(* Logix 5000 project; controller R400_500_XLS vendor 1 type 14 code 216 rev 31.11; software revision 31.01; part 10 of 32 *)
(* tags used below, declared in another part *)
   Alarm : SINT;   // Wait 3 seconds
   Cycles : UDT_CYCLE[11];
   DrnSmp : DINT;
   FC23_BaseConductivity : REAL;   // Base conductivity of the water prior to the injection
   Fill_Sump : DINT;
   M : DINT[5];   // Memory Bits
   MaxPressRecord : REAL;
   MinPressRecord : REAL;
   PureWaterTankFilling : BOOL;   // Start PWT filling
   Run : DINT;
   Service : DINT[2];   // Unused Service Mode Memory Bit
   Tmr : TIMER[107];
   WSH41_Hour : DINT;
   WSH41_Minute : DINT;
   WSH41_Second : DINT;
   abCycleDataToSCADA : BOOL[32];
   abInputToSCADA : BOOL[32];
   abOutputToSCADA : BOOL[32];
   aiCycleDataToSCADA : INT[16];
   AlarmTrigger : INT;   // Triggers the alarm screen if different of 0
   arAnalogInputToSCADA : REAL[8];
   arCycleDataToSCADA : REAL[8];
   bPureWaterFillingAuthorization : BOOL;   // Pure Water Filling Authorization Signal
   ChemCond : REAL;
   CR2Mode : SINT;   // 0= Cycle complete dry contact 1= External pure water valve
   CycleCounter : DINT;
   CyclePtr : DINT;   // Cycle Pointeur
   DryTemp : REAL;
   FinalRinseCond : REAL;
   I_Chm_1_Lvl_Sw : BOOL;   // Chemical Pump #1 level switch
   I_Chm_2_Lvl_Sw : BOOL;   // Chemical Pump #2 level switch
   I_Chm_3_Lvl_Sw : BOOL;   // Chemical Pump #3 level switch
   I_Chm_4_Lvl_Sw : BOOL;   // Chemical Pump #4 level switch
   I_Ld_Dr_Cls_Sw : BOOL;   // Load door close
   I_Ld_Dr_Obs_Sw : BOOL;   // Load door obstruction switch
   I_MCR : BOOL;   // MCR input
   I_Mtr_Ovrld : BOOL;   // Motor overload
   I_Pure_Water_Filling_Auth : BOOL;
   I_Pw_Tnk_Lvl_Sw : BOOL;   // Pure water tank level switch
   I_Pw_Tnk_Sft_Lvl_Sw : BOOL;   // Pure water tank safety level switch
   I_Shlf_Sw : BOOL;   // Shelf switch
   I_Smp_Lvl_Hgh : BOOL;   // Sump high level switch
   I_Smp_Lvl_Lw : BOOL;   // Sump low level switch
   I_Smp_Sft_Lvl_Sw : BOOL;   // Sump safety level switch
   I_Unld_Dr_Cls_Sw : BOOL;   // Unload door close
   I_Unld_Dr_Obs_Sw : BOOL;   // Unload door obstruction switch
   I_UnldDr_ClseSlnce_Bttn : BOOL;   // Door Close/ Silence button Unload Side
   I_UnldDr_Opn_Bttn : BOOL;   // Door Open button Unload side
   iAlarmToSCADA : INT;
   iSCADACycleCompleteTimeHr : INT;
   iSCADACycleCompleteTimeMin : INT;
   iSCADACycleCompleteTimeSec : INT;
   ONS_SCADA : INT;
   PmpPres : REAL;
   PureWaterTankFillingRequest : BOOL;
   PureWaterTankTemp : REAL;   // Pure water tank temperature
   Q_Adble_Alrm : BOOL;   // Audible Alarm and /Pilot Light: red connection
   Q_Chm_1 : BOOL;   // Chemical pump #1
   Q_Chm_2 : BOOL;   // Chemical pump #2
   Q_Chm_3 : BOOL;   // Chemical pump #3
   Q_Chm_4 : BOOL;   // Chemical pump #4
   Q_Cld_Wtr_Fll_Vlve : BOOL;   // Cold water sump fill valve
   Q_Cmmn_Alrm : BOOL;   // Dry contact For Alarm
   Q_Cndsr_Hflw_Vlve : BOOL;   // Condenser high flow cold water valve
   Q_Cndsr_Lflw_Vlve : BOOL;   // Condenser low flow cold water valve
   Q_Condensate_Return_Vlve : BOOL;   // Condensate Return CoolDown water valve
   Q_Cyc_Comp : BOOL;   // Dry Contact For Cycle Completed or Pure Water fill valve
   Q_Cyc_Run : BOOL;   // Pilot light: Green connection
   Q_Drn_Cldwn_Vlve : BOOL;   // Drain cool down water valve
   Q_Dry_Fan : BOOL;   // Vapor removal fan / Drying fan
   Q_Dry_Htr : BOOL;   // Drying heating elements
   Q_Dry_Iso_Vlve : BOOL;   // Drying Isolation Valve (Normally Closed Valve)
   Q_Ht_Rcvry_Tnk_Drn_Vlve : BOOL;   // Heat recovery tank drian valve
   Q_Ht_Wtr_Fll_Vlve : BOOL;   // Hot water sump fill valve
   Q_Int_Lght : BOOL;   // Interior Light
   Q_Ld_Dr_Clse_Vlv : BOOL;   // Load door close pilot valve
   Q_Ld_Dr_Opn_Vlv : BOOL;   // Load door open pilot valve
   Q_Pmp_Hgh_Spd : BOOL;   // Pump high speed
   Q_Pmp_Lw_Spd : BOOL;   // Pump low speed
   Q_Pure_Water_Filling_Request : BOOL;   // Pure Water Filling Request
   Q_Pw_Fll_Vlve : BOOL;   // Pure water sump/ Tank fill valve
   Q_Pw_Otlt_Vlve : BOOL;   // Pure water tank outlet valve
   Q_Pw_Tnk_Stm_Vlve : BOOL;   // PWT Steam Valve / Electric Heater
   Q_Smp_drn_Vlve : BOOL;   // Sump drain valve (Normally open valve)
   Q_Smp_Stm_Vlve : BOOL;   // Sump steam valve/ Electrical Heater
   Q_Trsfr_Vlve : BOOL;   // Transfer Valve (Normally Open Valve)
   Q_Unld_Dr_Clse_Vlve : BOOL;   // Unload door close pilot valve
   Q_Unld_Dr_Opn_Vlve : BOOL;   // Unload door open pilot valve
   rSCADACompensatedSetPoint : REAL;
   SumpTemp : REAL;   // Sump temperature in °C
   TreatmentPtr : DINT;
   udtPureWaterHandshakeFromSCADA : UDT_PORT_HANDSHAKE_FROM_SCADA;
   udtPureWaterHandshakeToSCADA : UDT_PORT_HANDSHAKE_TO_SCADA;
   Unit : Hrdwre;   // Unit Configuration
(* MainProgram, continued *)

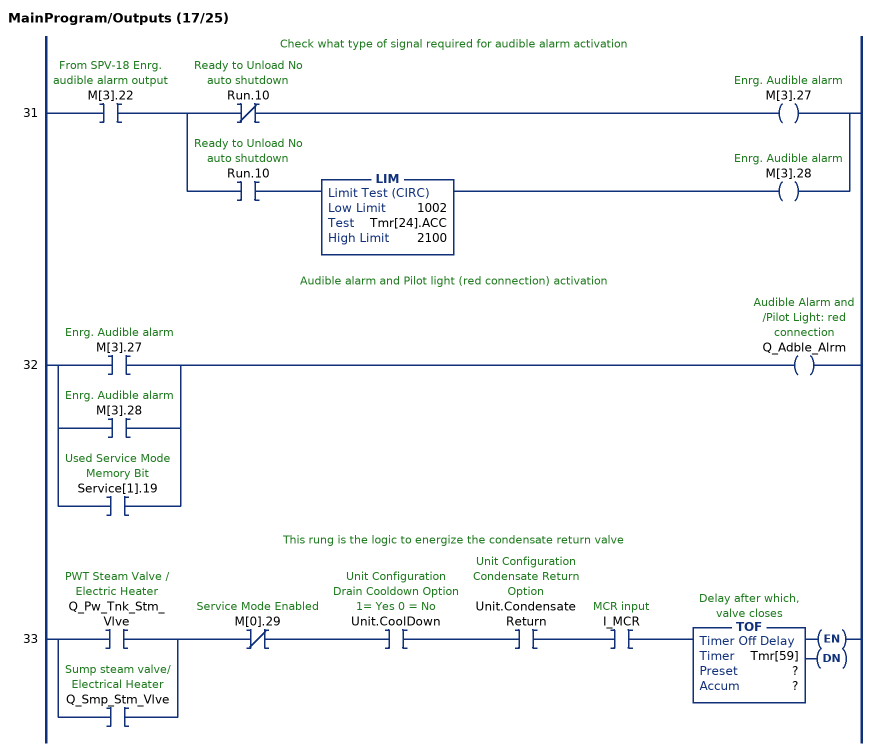
   [picture p153: MainProgram/Outputs rungs 31-33]
   // Check what type of signal required for audible alarm activation
   31: XIC(M[3].22)[XIO(Run.10) OTE(M[3].27) ,XIC(Run.10) LIM(1002,Tmr[24].ACC,2100) OTE(M[3].28) ];
   // Audible alarm and Pilot light (red connection) activation
   32: [XIC(M[3].27) ,XIC(M[3].28) ,XIC(Service[1].19) ]OTE(Q_Adble_Alrm);
   // This rung is the logic to energize the condensate return valve
   33: [XIC(Q_Pw_Tnk_Stm_Vlve) ,XIC(Q_Smp_Stm_Vlve) ]XIO(M[0].29)XIC(Unit.CoolDown)XIC(Unit.CondensateReturn)XIC(I_MCR)TOF(Tmr[59],?,?);
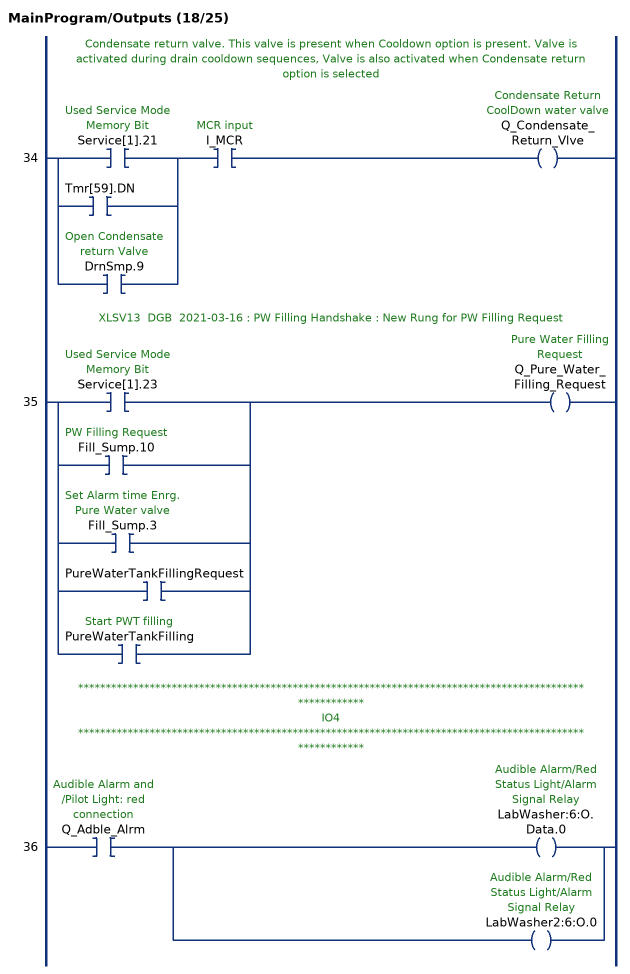
   // Condensate return valve. This valve is present when Cooldown option is present. Valve is activated during drain cooldown sequences, Valve is also activated when Condensate return option is selected
   34: [XIC(Service[1].21) ,XIC(Tmr[59].DN) ,XIC(DrnSmp.9) ]XIC(I_MCR)OTE(Q_Condensate_Return_Vlve);
   // XLSV13  DGB  2021-03-16 : PW Filling Handshake : New Rung for PW Filling Request
   35: [XIC(Service[1].23) ,XIC(Fill_Sump.10) ,XIC(Fill_Sump.3) ,XIC(PureWaterTankFillingRequest) ,XIC(PureWaterTankFilling) ]OTE(Q_Pure_Water_Filling_Request);
   // ********************************************************************************************************
   // IO4
   // ********************************************************************************************************
   36: XIC(Q_Adble_Alrm)[OTE(LabWasher:6:O.Data.0) ,OTE(LabWasher2:6:O.0) ];
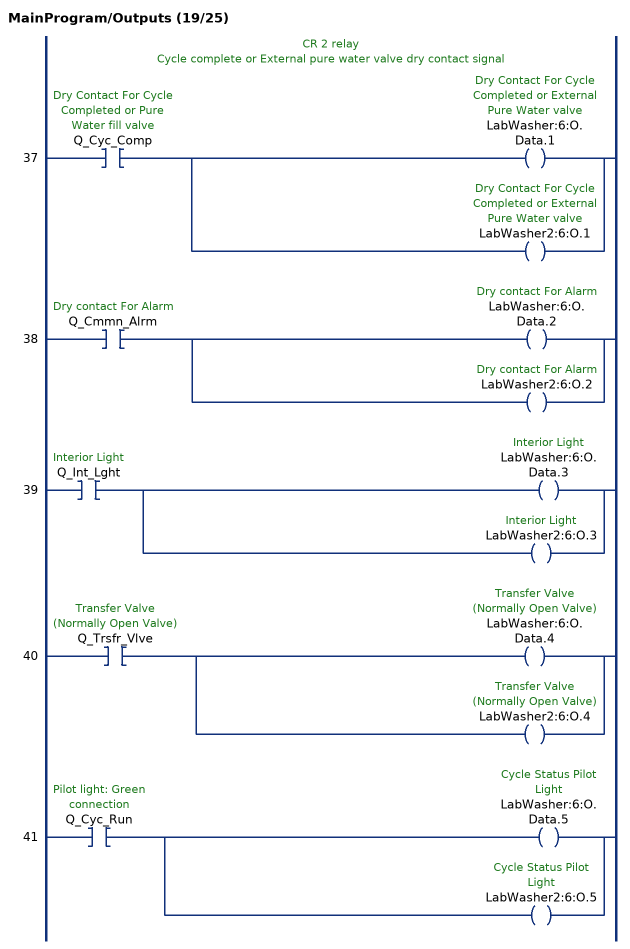
   // CR 2 relay
   // Cycle complete or External pure water valve dry contact signal
   37: XIC(Q_Cyc_Comp)[OTE(LabWasher:6:O.Data.1) ,OTE(LabWasher2:6:O.1) ];
   38: XIC(Q_Cmmn_Alrm)[OTE(LabWasher:6:O.Data.2) ,OTE(LabWasher2:6:O.2) ];
   39: XIC(Q_Int_Lght)[OTE(LabWasher:6:O.Data.3) ,OTE(LabWasher2:6:O.3) ];
   40: XIC(Q_Trsfr_Vlve)[OTE(LabWasher:6:O.Data.4) ,OTE(LabWasher2:6:O.4) ];
   41: XIC(Q_Cyc_Run)[OTE(LabWasher:6:O.Data.5) ,OTE(LabWasher2:6:O.5) ];
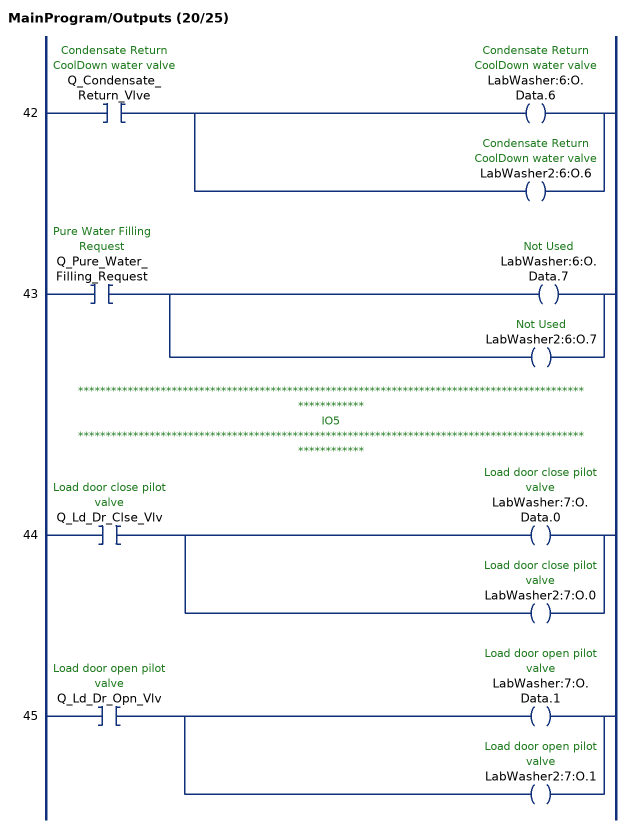
   42: XIC(Q_Condensate_Return_Vlve)[OTE(LabWasher:6:O.Data.6) ,OTE(LabWasher2:6:O.6) ];
   43: XIC(Q_Pure_Water_Filling_Request)[OTE(LabWasher:6:O.Data.7) ,OTE(LabWasher2:6:O.7) ];
   // ********************************************************************************************************
   // IO5
   // ********************************************************************************************************
   44: XIC(Q_Ld_Dr_Clse_Vlv)[OTE(LabWasher:7:O.Data.0) ,OTE(LabWasher2:7:O.0) ];
   45: XIC(Q_Ld_Dr_Opn_Vlv)[OTE(LabWasher:7:O.Data.1) ,OTE(LabWasher2:7:O.1) ];
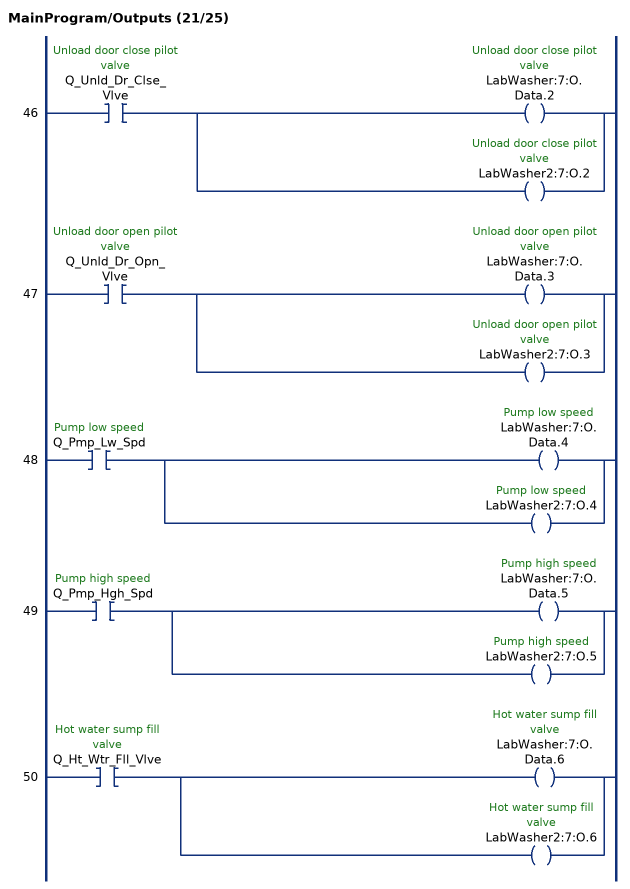
   46: XIC(Q_Unld_Dr_Clse_Vlve)[OTE(LabWasher:7:O.Data.2) ,OTE(LabWasher2:7:O.2) ];
   47: XIC(Q_Unld_Dr_Opn_Vlve)[OTE(LabWasher:7:O.Data.3) ,OTE(LabWasher2:7:O.3) ];
   48: XIC(Q_Pmp_Lw_Spd)[OTE(LabWasher:7:O.Data.4) ,OTE(LabWasher2:7:O.4) ];
   49: XIC(Q_Pmp_Hgh_Spd)[OTE(LabWasher:7:O.Data.5) ,OTE(LabWasher2:7:O.5) ];
   50: XIC(Q_Ht_Wtr_Fll_Vlve)[OTE(LabWasher:7:O.Data.6) ,OTE(LabWasher2:7:O.6) ];
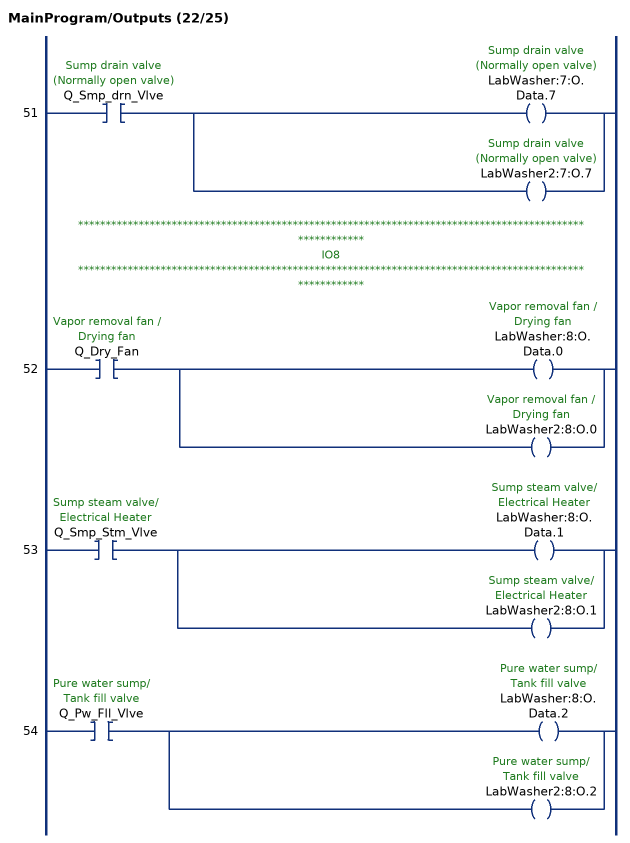
   51: XIC(Q_Smp_drn_Vlve)[OTE(LabWasher:7:O.Data.7) ,OTE(LabWasher2:7:O.7) ];
   // ********************************************************************************************************
   // IO8
   // ********************************************************************************************************
   52: XIC(Q_Dry_Fan)[OTE(LabWasher:8:O.Data.0) ,OTE(LabWasher2:8:O.0) ];
   53: XIC(Q_Smp_Stm_Vlve)[OTE(LabWasher:8:O.Data.1) ,OTE(LabWasher2:8:O.1) ];
   54: XIC(Q_Pw_Fll_Vlve)[OTE(LabWasher:8:O.Data.2) ,OTE(LabWasher2:8:O.2) ];
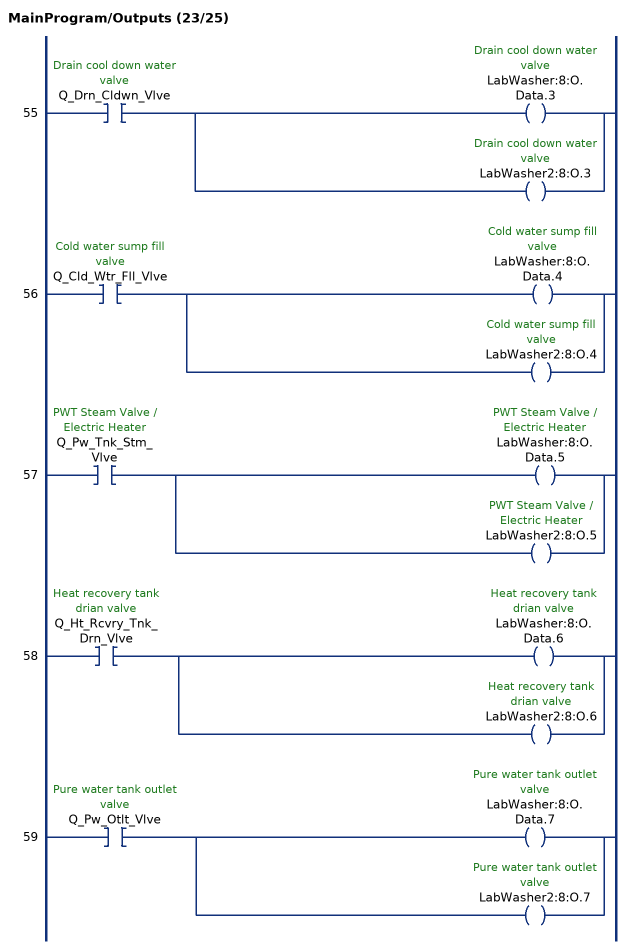
   55: XIC(Q_Drn_Cldwn_Vlve)[OTE(LabWasher:8:O.Data.3) ,OTE(LabWasher2:8:O.3) ];
   56: XIC(Q_Cld_Wtr_Fll_Vlve)[OTE(LabWasher:8:O.Data.4) ,OTE(LabWasher2:8:O.4) ];
   57: XIC(Q_Pw_Tnk_Stm_Vlve)[OTE(LabWasher:8:O.Data.5) ,OTE(LabWasher2:8:O.5) ];
   58: XIC(Q_Ht_Rcvry_Tnk_Drn_Vlve)[OTE(LabWasher:8:O.Data.6) ,OTE(LabWasher2:8:O.6) ];
   59: XIC(Q_Pw_Otlt_Vlve)[OTE(LabWasher:8:O.Data.7) ,OTE(LabWasher2:8:O.7) ];
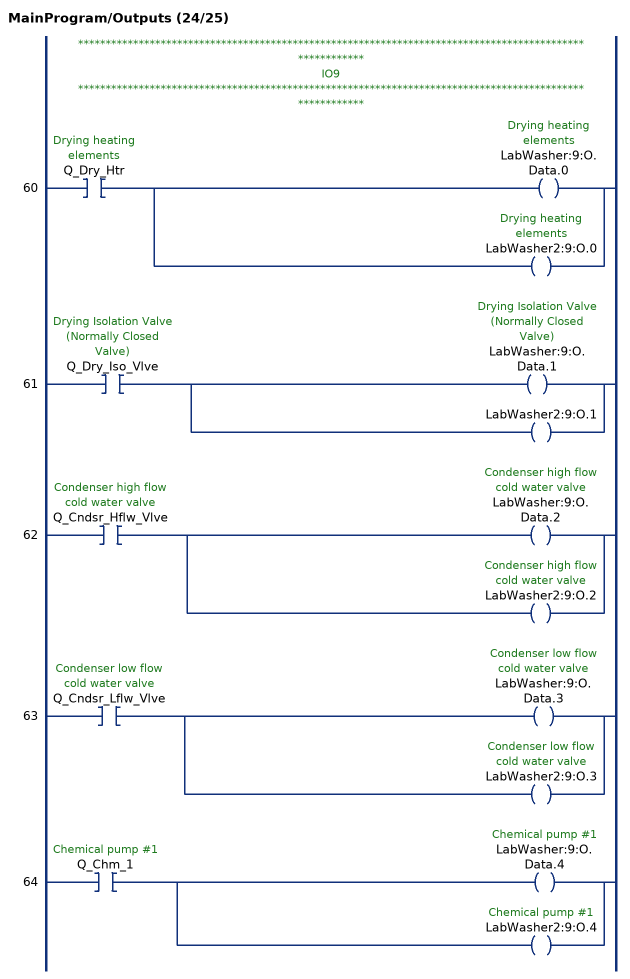
   // ********************************************************************************************************
   // IO9
   // ********************************************************************************************************
   60: XIC(Q_Dry_Htr)[OTE(LabWasher:9:O.Data.0) ,OTE(LabWasher2:9:O.0) ];
   61: XIC(Q_Dry_Iso_Vlve)[OTE(LabWasher:9:O.Data.1) ,OTE(LabWasher2:9:O.1) ];
   62: XIC(Q_Cndsr_Hflw_Vlve)[OTE(LabWasher:9:O.Data.2) ,OTE(LabWasher2:9:O.2) ];
   63: XIC(Q_Cndsr_Lflw_Vlve)[OTE(LabWasher:9:O.Data.3) ,OTE(LabWasher2:9:O.3) ];
   64: XIC(Q_Chm_1)[OTE(LabWasher:9:O.Data.4) ,OTE(LabWasher2:9:O.4) ];
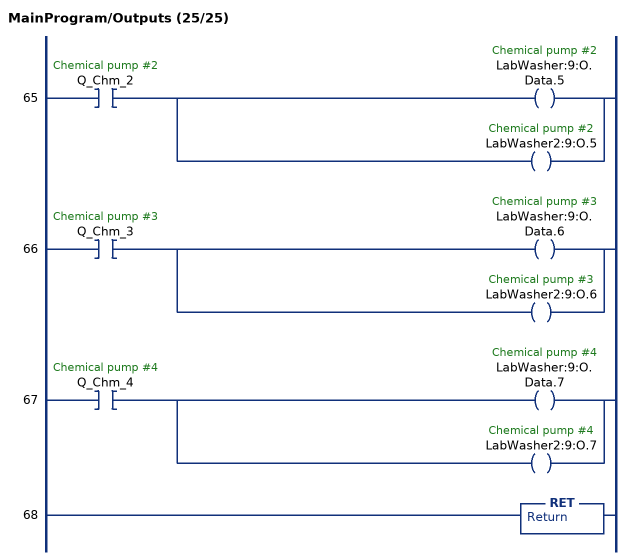
   65: XIC(Q_Chm_2)[OTE(LabWasher:9:O.Data.5) ,OTE(LabWasher2:9:O.5) ];
   66: XIC(Q_Chm_3)[OTE(LabWasher:9:O.Data.6) ,OTE(LabWasher2:9:O.6) ];
   67: XIC(Q_Chm_4)[OTE(LabWasher:9:O.Data.7) ,OTE(LabWasher2:9:O.7) ];
   68: RET();
END_ROUTINE

ROUTINE SCADA   (* ladder *)
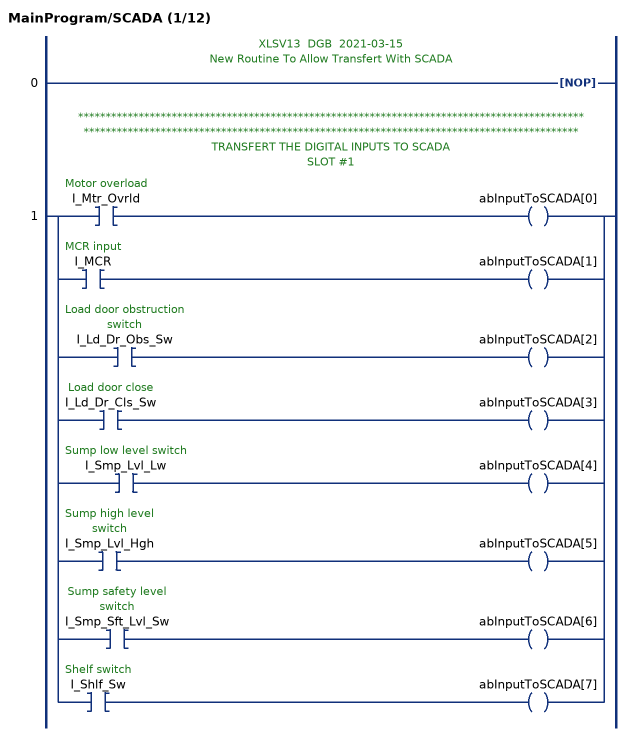
   // XLSV13  DGB  2021-03-15
   // New Routine To Allow Transfert With SCADA
   0: NOP();
   // **************************************************************************************************************************************************************************************
   // TRANSFERT THE DIGITAL INPUTS TO SCADA
   // SLOT #1
   1: [XIC(I_Mtr_Ovrld) OTE(abInputToSCADA[0]) ,XIC(I_MCR) OTE(abInputToSCADA[1]) ,XIC(I_Ld_Dr_Obs_Sw) OTE(abInputToSCADA[2]) ,XIC(I_Ld_Dr_Cls_Sw) OTE(abInputToSCADA[3]) ,XIC(I_Smp_Lvl_Lw) OTE(abInputToSCADA[4]) ,XIC(I_Smp_Lvl_Hgh) OTE(abInputToSCADA[5]) ,XIC(I_Smp_Sft_Lvl_Sw) OTE(abInputToSCADA[6]) ,XIC(I_Shlf_Sw) OTE(abInputToSCADA[7]) ];
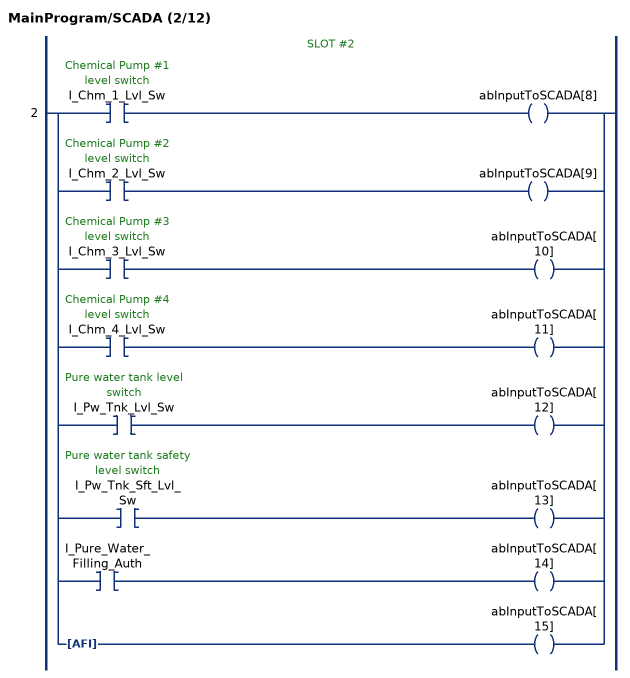
   // SLOT #2
   2: [XIC(I_Chm_1_Lvl_Sw) OTE(abInputToSCADA[8]) ,XIC(I_Chm_2_Lvl_Sw) OTE(abInputToSCADA[9]) ,XIC(I_Chm_3_Lvl_Sw) OTE(abInputToSCADA[10]) ,XIC(I_Chm_4_Lvl_Sw) OTE(abInputToSCADA[11]) ,XIC(I_Pw_Tnk_Lvl_Sw) OTE(abInputToSCADA[12]) ,XIC(I_Pw_Tnk_Sft_Lvl_Sw) OTE(abInputToSCADA[13]) ,XIC(I_Pure_Water_Filling_Auth) OTE(abInputToSCADA[14]) ,AFI() OTE(abInputToSCADA[15]) ];
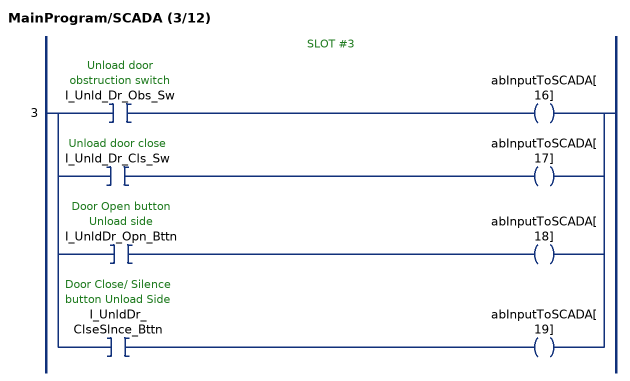
   // SLOT #3
   3: [XIC(I_Unld_Dr_Obs_Sw) OTE(abInputToSCADA[16]) ,XIC(I_Unld_Dr_Cls_Sw) OTE(abInputToSCADA[17]) ,XIC(I_UnldDr_Opn_Bttn) OTE(abInputToSCADA[18]) ,XIC(I_UnldDr_ClseSlnce_Bttn) OTE(abInputToSCADA[19]) ];
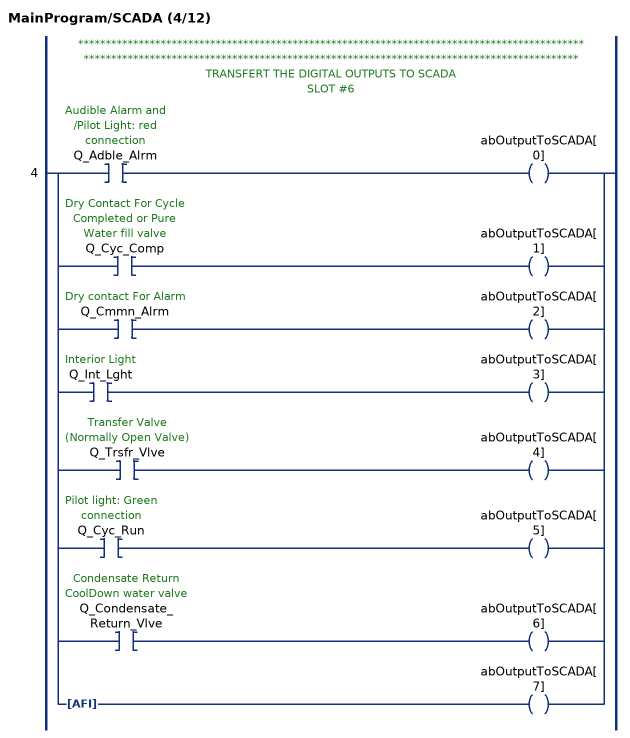
   // **************************************************************************************************************************************************************************************
   // TRANSFERT THE DIGITAL OUTPUTS TO SCADA
   // SLOT #6
   4: [XIC(Q_Adble_Alrm) OTE(abOutputToSCADA[0]) ,XIC(Q_Cyc_Comp) OTE(abOutputToSCADA[1]) ,XIC(Q_Cmmn_Alrm) OTE(abOutputToSCADA[2]) ,XIC(Q_Int_Lght) OTE(abOutputToSCADA[3]) ,XIC(Q_Trsfr_Vlve) OTE(abOutputToSCADA[4]) ,XIC(Q_Cyc_Run) OTE(abOutputToSCADA[5]) ,XIC(Q_Condensate_Return_Vlve) OTE(abOutputToSCADA[6]) ,AFI() OTE(abOutputToSCADA[7]) ];
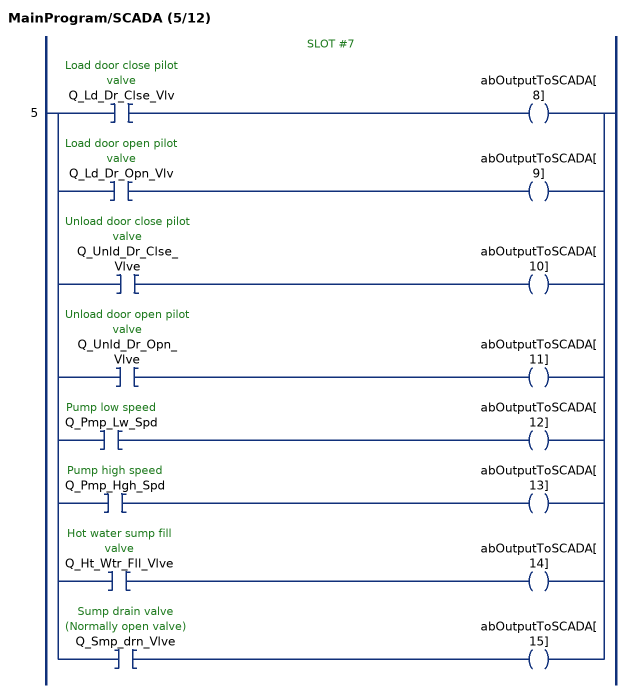
   // SLOT #7
   5: [XIC(Q_Ld_Dr_Clse_Vlv) OTE(abOutputToSCADA[8]) ,XIC(Q_Ld_Dr_Opn_Vlv) OTE(abOutputToSCADA[9]) ,XIC(Q_Unld_Dr_Clse_Vlve) OTE(abOutputToSCADA[10]) ,XIC(Q_Unld_Dr_Opn_Vlve) OTE(abOutputToSCADA[11]) ,XIC(Q_Pmp_Lw_Spd) OTE(abOutputToSCADA[12]) ,XIC(Q_Pmp_Hgh_Spd) OTE(abOutputToSCADA[13]) ,XIC(Q_Ht_Wtr_Fll_Vlve) OTE(abOutputToSCADA[14]) ,XIC(Q_Smp_drn_Vlve) OTE(abOutputToSCADA[15]) ];
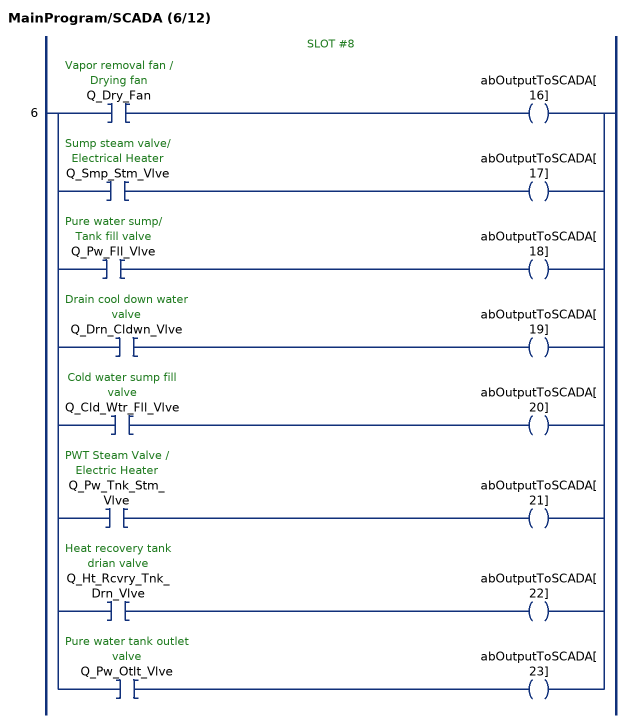
   // SLOT #8
   6: [XIC(Q_Dry_Fan) OTE(abOutputToSCADA[16]) ,XIC(Q_Smp_Stm_Vlve) OTE(abOutputToSCADA[17]) ,XIC(Q_Pw_Fll_Vlve) OTE(abOutputToSCADA[18]) ,XIC(Q_Drn_Cldwn_Vlve) OTE(abOutputToSCADA[19]) ,XIC(Q_Cld_Wtr_Fll_Vlve) OTE(abOutputToSCADA[20]) ,XIC(Q_Pw_Tnk_Stm_Vlve) OTE(abOutputToSCADA[21]) ,XIC(Q_Ht_Rcvry_Tnk_Drn_Vlve) OTE(abOutputToSCADA[22]) ,XIC(Q_Pw_Otlt_Vlve) OTE(abOutputToSCADA[23]) ];
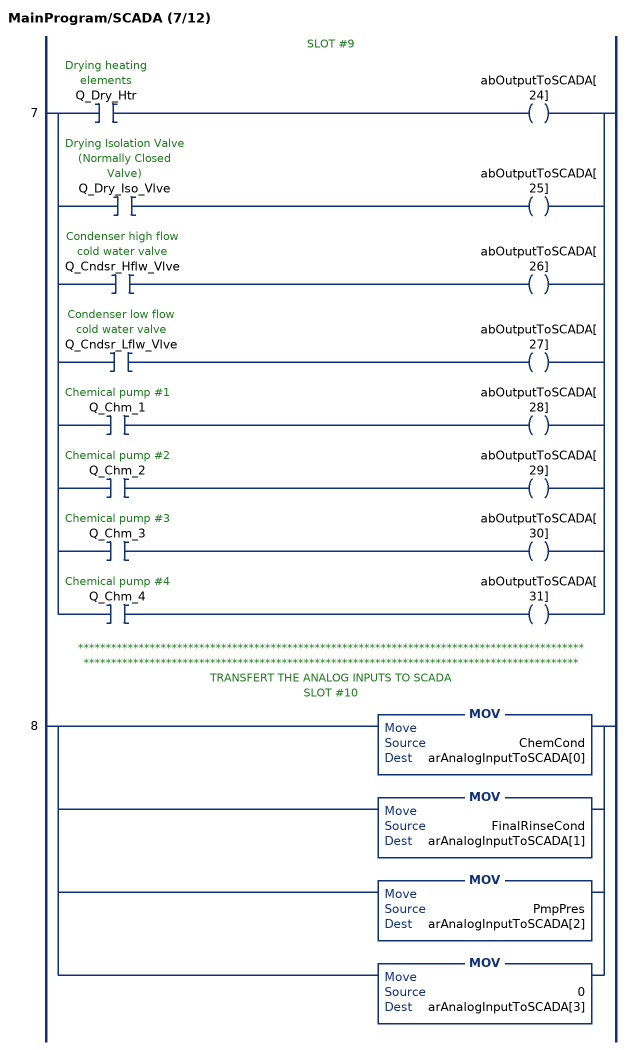
   // SLOT #9
   7: [XIC(Q_Dry_Htr) OTE(abOutputToSCADA[24]) ,XIC(Q_Dry_Iso_Vlve) OTE(abOutputToSCADA[25]) ,XIC(Q_Cndsr_Hflw_Vlve) OTE(abOutputToSCADA[26]) ,XIC(Q_Cndsr_Lflw_Vlve) OTE(abOutputToSCADA[27]) ,XIC(Q_Chm_1) OTE(abOutputToSCADA[28]) ,XIC(Q_Chm_2) OTE(abOutputToSCADA[29]) ,XIC(Q_Chm_3) OTE(abOutputToSCADA[30]) ,XIC(Q_Chm_4) OTE(abOutputToSCADA[31]) ];
   // **************************************************************************************************************************************************************************************
   // TRANSFERT THE ANALOG INPUTS TO SCADA
   // SLOT #10
   8: [MOV(ChemCond,arAnalogInputToSCADA[0]) ,MOV(FinalRinseCond,arAnalogInputToSCADA[1]) ,MOV(PmpPres,arAnalogInputToSCADA[2]) ,MOV(0,arAnalogInputToSCADA[3]) ];
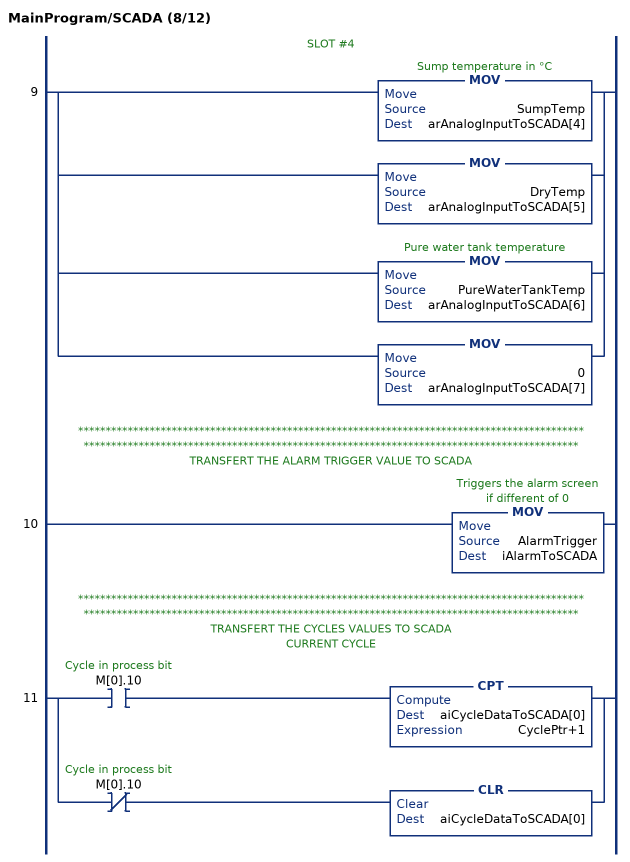
   // SLOT #4
   9: [MOV(SumpTemp,arAnalogInputToSCADA[4]) ,MOV(DryTemp,arAnalogInputToSCADA[5]) ,MOV(PureWaterTankTemp,arAnalogInputToSCADA[6]) ,MOV(0,arAnalogInputToSCADA[7]) ];
   // **************************************************************************************************************************************************************************************
   // TRANSFERT THE ALARM TRIGGER VALUE TO SCADA
   10: MOV(AlarmTrigger,iAlarmToSCADA);
   // **************************************************************************************************************************************************************************************
   // TRANSFERT THE CYCLES VALUES TO SCADA
   // CURRENT CYCLE
   11: [XIC(M[0].10) CPT(aiCycleDataToSCADA[0],CyclePtr+1) ,XIO(M[0].10) CLR(aiCycleDataToSCADA[0]) ];
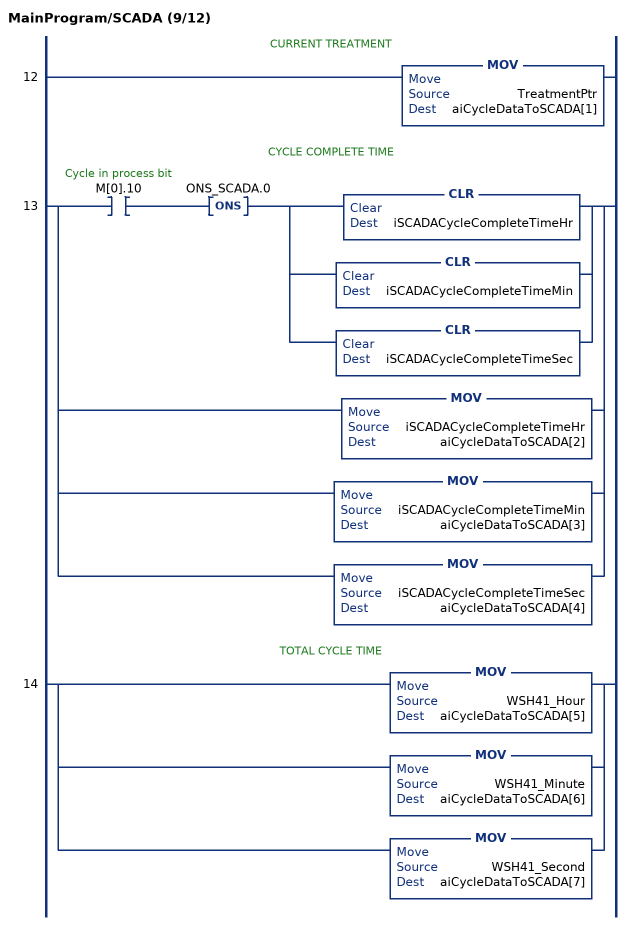
   // CURRENT TREATMENT
   12: MOV(TreatmentPtr,aiCycleDataToSCADA[1]);
   // CYCLE COMPLETE TIME
   13: [XIC(M[0].10) ONS(ONS_SCADA.0) [CLR(iSCADACycleCompleteTimeHr) ,CLR(iSCADACycleCompleteTimeMin) ,CLR(iSCADACycleCompleteTimeSec) ] ,MOV(iSCADACycleCompleteTimeHr,aiCycleDataToSCADA[2]) ,MOV(iSCADACycleCompleteTimeMin,aiCycleDataToSCADA[3]) ,MOV(iSCADACycleCompleteTimeSec,aiCycleDataToSCADA[4]) ];
   // TOTAL CYCLE TIME
   14: [MOV(WSH41_Hour,aiCycleDataToSCADA[5]) ,MOV(WSH41_Minute,aiCycleDataToSCADA[6]) ,MOV(WSH41_Second,aiCycleDataToSCADA[7]) ];
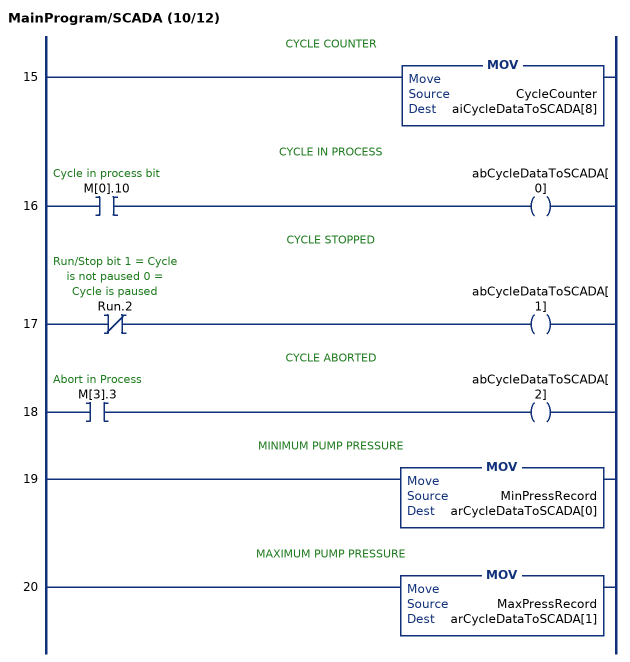
   // CYCLE COUNTER
   15: MOV(CycleCounter,aiCycleDataToSCADA[8]);
   // CYCLE IN PROCESS
   16: XIC(M[0].10)OTE(abCycleDataToSCADA[0]);
   // CYCLE STOPPED
   17: XIO(Run.2)OTE(abCycleDataToSCADA[1]);
   // CYCLE ABORTED
   18: XIC(M[3].3)OTE(abCycleDataToSCADA[2]);
   // MINIMUM PUMP PRESSURE
   19: MOV(MinPressRecord,arCycleDataToSCADA[0]);
   // MAXIMUM PUMP PRESSURE
   20: MOV(MaxPressRecord,arCycleDataToSCADA[1]);
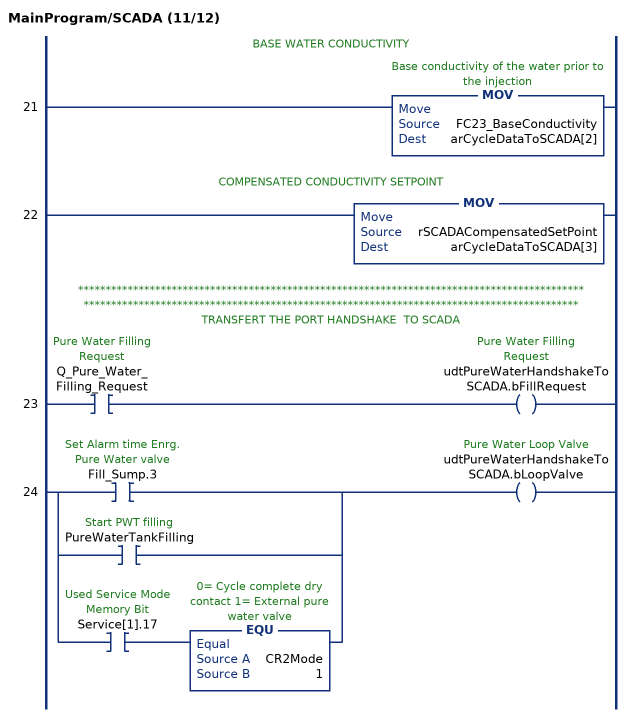
   // BASE WATER CONDUCTIVITY
   21: MOV(FC23_BaseConductivity,arCycleDataToSCADA[2]);
   // COMPENSATED CONDUCTIVITY SETPOINT
   22: MOV(rSCADACompensatedSetPoint,arCycleDataToSCADA[3]);
   // **************************************************************************************************************************************************************************************
   // TRANSFERT THE PORT HANDSHAKE  TO SCADA
   23: XIC(Q_Pure_Water_Filling_Request)OTE(udtPureWaterHandshakeToSCADA.bFillRequest);
   24: [XIC(Fill_Sump.3) ,XIC(PureWaterTankFilling) ,XIC(Service[1].17) EQU(CR2Mode,1) ]OTE(udtPureWaterHandshakeToSCADA.bLoopValve);
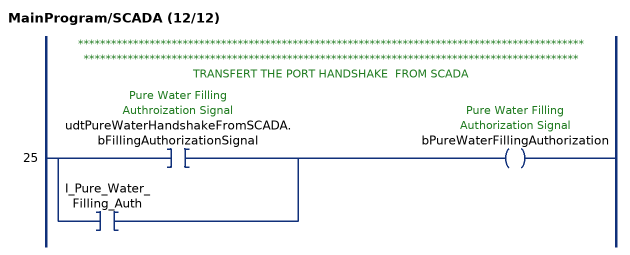
   // **************************************************************************************************************************************************************************************
   // TRANSFERT THE PORT HANDSHAKE  FROM SCADA
   25: [XIC(udtPureWaterHandshakeFromSCADA.bFillingAuthorizationSignal) ,XIC(I_Pure_Water_Filling_Auth) ]OTE(bPureWaterFillingAuthorization);
END_ROUTINE
